Fanuc TP program (LS listing): PrecPr.LS

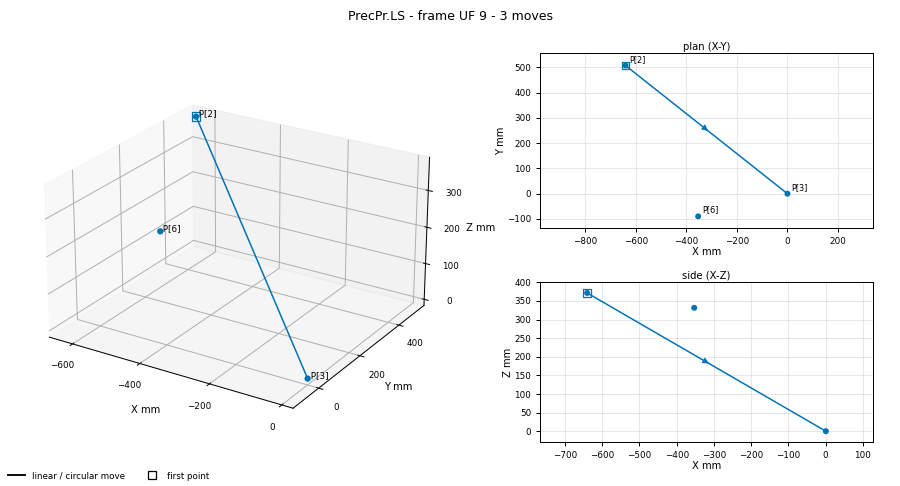
[picture p0: tool path of PrecPr.LS in frame UF 9, 3 of 6 moves have a stored position in this frame; points joined in program order, loops and branches not executed]
/PROG  PrecPr
/ATTR
OWNER		= MNEDITOR;
COMMENT		= "RoboDK sequence";
PROG_SIZE	= 0;
CREATE		= DATE 31-12-14  TIME 12:00:00;
MODIFIED	= DATE 31-12-14  TIME 12:00:00;
FILE_NAME	= PrecPr;
VERSION		= 0;
LINE_COUNT	= 27;
MEMORY_SIZE	= 0;
PROTECT		= READ_WRITE;
TCD:  STACK_SIZE	= 0,
      TASK_PRIORITY	= 50,
      TIME_SLICE	= 0,
      BUSY_LAMP_OFF	= 0,
      ABORT_REQUEST	= 0,
      PAUSE_REQUEST	= 0;
DEFAULT_GROUP	= 1,*,*,*,*;
CONTROL_CODE	= 00000000 00000000;
/MN
   1:  ! Program generated by RoboDK v6.0.7 for Fanuc M-1iA/0.5S on XX ;
   2:  ! /XX/XXXX 18:00:00 ;
   3:  ! Using nominal kinematics. ;
   4:  PR[9,1]=0.000 ;
   5:  PR[9,2]=-0.001 ;
   6:  PR[9,3]=1000.000 ;
   7:  PR[9,4]=90.000 ;
   8:  PR[9,5]=-0.500 ;
   9:  PR[9,6]=0.123 ;
  10:  UFRAME[9]=PR[9] ;
  11:  UFRAME_NUM=9 ;
  12:  PR[9,1]=0.125 ;
  13:  PR[9,2]=-0.375 ;
  14:  PR[9,3]=123.457 ;
  15:  PR[9,4]=-45.250 ;
  16:  PR[9,5]=0.000 ;
  17:  PR[9,6]=0.000 ;
  18:  UTOOL[9]=PR[9] ;
  19:  UTOOL_NUM=9 ;
  20:J P[1] 20% FINE ;
  21:L P[2] 200mm/sec FINE ;
  22:L P[3] 200mm/sec FINE ;
  23:J P[4] 20% FINE ;
  24:J P[5] 20% FINE ;
  25:  WAIT  0.00(sec) ;
  26:  WAIT  1.00(sec) ;
  27:L P[6] 67mm/sec FINE ;
/POS
P[1]{
   GP1:
    UF : 9, UT : 9,
	J1=    12.345600 deg,	J2=    -45.678900 deg,	J3=    78.901300  mm,
	J4=    -0.500000 deg
};
P[2]{
   GP1:
    UF : 9, UT : 9,        CONFIG : 'L, 0, 0, 0',
	X =  -640.585  mm,	Y =   506.981  mm,	Z =   371.534  mm,
	W =  -165.500 deg,	P =    50.000 deg,	R =   150.000 deg
};
P[3]{
   GP1:
    UF : 9, UT : 9,        CONFIG : 'L, 0, 0, 0',
	X =     0.500  mm,	Y =    -0.500  mm,	Z =     0.250  mm,
	W =   180.000 deg,	P =    -0.005 deg,	R =     0.005 deg
};
P[4]{
   GP1:
    UF : 9, UT : 9,
	J1=    -12.345400 deg,	J2=    45.678500 deg,	J3=    -78.900000  mm,
	J4=    0.500000 deg
};
P[5]{
   GP1:
    UF : 9, UT : 9,
	J1=    -12.345400 deg,	J2=    45.678500 deg,	J3=    -78.900000  mm,
	J4=    0.500000 deg
};
P[6]{
   GP1:
    UF : 9, UT : 9,        CONFIG : 'L, 0, 0, 0',
	X =  -353.026  mm,	Y =   -90.135  mm,	Z =   331.702  mm,
	W =  -169.444 deg,	P =    40.650 deg,	R =   178.023 deg
};
/END
